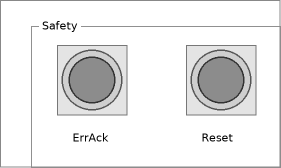
VISUALIZATION Safety  // 281x168
    GroupBox (31,18 250x150), "Safety"
        PushSwitchLed (155,27 70x70), variable: GVL_Safety.Restart, behaviour: TOGGLE, style: Switch-PushSwitchLed-Gray
        PushSwitchLed (26,27 70x70), variable: GVL_Safety.ErrAck, behaviour: TOGGLE, style: Switch-PushSwitchLed-Gray
        Label (21,105 77x30), "ErrAck"
        Label (157,105 59x30), "Reset"
END_VISUALIZATION

(* stored: Version 1.1.0.1, ProductVersion 3.1.4024.15
   Visu Safety: Id {e4c18a57-4875-4f76-96ba-a974204b1731} *)
